FUNCTION_BLOCK FB_Auswerfer
VAR_INPUT
END_VAR
VAR_OUTPUT
END_VAR
VAR
END_VAR

GVL_IO.xVentilAuswerferAS := GVL_IO.xWeicheRejectBereit;
GVL_IO.xVentilAuswerferGS := NOT GVL_IO.xWeicheRejectBereit;

GVL_IO.xAuswerferBereit := GVL_IO.xZylinderAuswerferAS;

END_FUNCTION_BLOCK

(* stored: Version 1.1.0.1
   POU FB_Auswerfer: Id {f5fe8941-58c6-4719-9129-89b405f01ed3}, SpecialFunc None *)
